(* IEC 61131-3 sources: Caravan/Archiv/12-04-19/Stations/Terminal/HMI/Network/STDSettingsHMI, 1 file *)

(* ---- ONE_STDSettingsHMI_Table.st ---- *)
#define OBJECTS_CONFIG

//Define part of class ProjectGlobal
// Eigenschaften der Bildschirm-Informationen
//----------------------------------------------------------------------------------
#define Global_NumScreenInfos                            100                                 // Anzahl der reservierten Einträge für die Bildschirminformation

#define Global_MenueScreenNr                             10                                  // Bildschirm-Nummer des Menüs (Startseite)

#define Global_MenueMin                                  5                                   // Bildschirm-Nummer Alarme(*Ez0999*)

#define Global_MenueMax                                  4410                                // Bildschirm-Nummer Login Screens(*Ez0999*)

#define PRJGLOBAL_MAX_STATION                            255                                 // Highest possible LSE Station-Number

#define PRJGLOBAL_STATION_INTERN                         0                                   // Identifier for internal LSE-Station

#define PRJGLOBAL_STATION_EXTERN                         1                                   // Identifier for TCPIP1 LSE-Station

#define     CMD_GETIPOverStation      1000
//Define part of class USBDetection
#define USB_StringLength                              _strlen("C:\")          // Länge des Strings für das aktuelle Laufwerk

FUNCTION GLOBAL TAB ONE_STDSettingsHMI
-1$UINT, 0$UINT,
2$UINT, 0$UINT,

9$UDINT,
TO_UDINT(3788417926), "_Global", 0$UINT, 14$UINT, 0$UINT,
TO_UDINT(3877617373), "_SyncTimeHMI", 2$UINT, 0$UINT, 1$UINT,
TO_UDINT(2225119864), "MerkerEx", 1$UINT, 21$UINT, 1$UINT,
TO_UDINT(1462004836), "ProjectGlobal", 1$UINT, 16$UINT, 1$UINT,
TO_UDINT(1903583397), "Ram", 1$UINT, 3$UINT, 2$UINT,
TO_UDINT(1850111279), "String", 1$UINT, 10$UINT, 1$UINT,
TO_UDINT(2898603620), "StringInternal", 1$UINT, 82$UINT, 0$UINT,
TO_UDINT(216038476), "USBDetection", 1$UINT, 5$UINT, 1$UINT,
TO_UDINT(3232495061), "VirtualBaseInit", 1$UINT, 3$UINT, 0$UINT,

_NO_ATTR, TO_UDINT(3114404899), "SYNCTIMEHMI",

1$UINT, TO_UDINT(1839314391), "USBDETECTION1\USBDRIVELETTER\MERKEREX0",

_NO_ATTR, TO_UDINT(2925151108), "GLOBALSCREEN1",

1$UINT, TO_UDINT(2793771928), "GLOBALSCREEN1\OFFDATE",
1$UINT, TO_UDINT(1670331559), "GLOBALSCREEN1\OFFTIME",

1$UINT, TO_UDINT(267725679), "USBDETECTION1\USBDRIVELETTER",

_NO_ATTR, TO_UDINT(4240048752), "USBDETECTION1",

//Internal connections
0$UDINT,
4$UDINT,
TO_UDINT(2), "OffDate", TO_UDINT(3),
TO_UDINT(2), "OffTime", TO_UDINT(4),
TO_UDINT(5), "MerkerEx0", TO_UDINT(1),
TO_UDINT(6), "USBDriveLetter", TO_UDINT(5),
0$UDINT,
1$UDINT,
TO_UDINT(5), "DataBuffer", TO_UDINT(1), "m_udLength",

//Initialization values
0$UDINT,
5$UDINT,
TO_UDINT(1), "ThreadSafe", TO_UDINT(0),//|STDSettingsHMI.USBDriveLetter\USBDetection1\MerkerEx0.ThreadSafe;
TO_UDINT(2), "OwnStationNumber", TO_UDINT(-1),//|STDSettingsHMI.GlobalScreen1.OwnStationNumber;
TO_UDINT(2), "ExtStationNumber", TO_UDINT(-1),//|STDSettingsHMI.GlobalScreen1.ExtStationNumber;
TO_UDINT(2), "ProjectReady", TO_UDINT(0),//|STDSettingsHMI.GlobalScreen1.ProjectReady;
TO_UDINT(5), "SingleRealloc", TO_UDINT(1),//|STDSettingsHMI.USBDetection1\USBDriveLetter.SingleRealloc;

//Symbolic initialization values
0$UDINT,
0$UDINT,

//Initialization of string values
0$UDINT,
0$UDINT,

//Configuration of tasks (RealTime, Cyclic, Background)
0$UDINT,
0$UDINT,

0$UDINT,
0$UDINT,

0$UDINT,
1$UDINT,
TO_UDINT(0), (100)$UDINT, 4194303$DINT, 	//SYNCTIMEHMI

//External connections
0$UDINT,
6$UDINT,
TO_UDINT(0), "ActDate", C_DIR, TO_UDINT(3035062039), "SysDateTime","SysDate",
TO_UDINT(0), "ActTime", C_DIR, TO_UDINT(3035062039), "SysDateTime","SysTime",
TO_UDINT(2), "Lse", C_DIR, TO_UDINT(299963966), "Lse","Lse",
TO_UDINT(2), "SysDate", C_DIR, TO_UDINT(3035062039), "SysDateTime","SysDate",
TO_UDINT(2), "SysTime", C_DIR, TO_UDINT(3035062039), "SysDateTime","SysTime",
TO_UDINT(6), "Lse", C_DIR, TO_UDINT(299963966), "Lse","Lse",

//Magic internal connections
0$UDINT,
0$UDINT,

//Configuration of timeslots of tasks (RealTime, Cyclic)
#ifdef __LSLLDR_TIMESLOTS__
0$UDINT,
0$UDINT,

0$UDINT,
0$UDINT,

#endif //__LSLLDR_TIMESLOTS__

//MultiMaster connections
#ifdef __LSLLDR_MULTIMASTER__
0$UDINT,
2$UDINT,
TO_UDINT(0), "SetDate", C_TRY, TO_UDINT(619908241), "MachineControl.SyncTimePLC.SyncDate",
TO_UDINT(0), "SetTime", C_TRY, TO_UDINT(3791233966), "MachineControl.SyncTimePLC.SyncTime",
#endif //__LSLLDR_MULTIMASTER__

//Configuration for task ID (RealTime, CyclicTime)
#ifdef __LSLLDR_TASKID__
"\\\\TASKS2  "
0$UDINT,
0$UDINT,

0$UDINT,
0$UDINT,

0$UDINT,
1$UDINT,
(0)$UDINT, 	//SYNCTIMEHMI

#endif //__LSLLDR_TASKID__

END_FUNCTION
